{attribute 'pack_mode' := '1'}
TYPE ST_BatPublishData :
STRUCT
	Header		:	ST_MqttHeader;
	Devices		:	ARRAY[0..GVL_PARAM.BMS_COUNT-1] OF ST_BatPublish_V1;
END_STRUCT
END_TYPE

(* stored: Version 1.1.0.1, ProductVersion 3.1.4024.15
   DUT ST_BatPublishData: Id {383c9f48-002c-4e4b-a147-9a11aad45ff3} *)
